FUNCTION_BLOCK PID_SAMPLE_COORDINATOR (* Experimental; offline checks only; native export/runtime pending *)
  (* Standard: 61499-2 *)
  (* Version 0.1, 2026-10-20, Guilherme *)
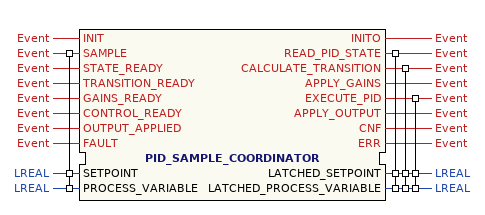
  EVENT_INPUT
    INIT;
    SAMPLE WITH SETPOINT, PROCESS_VARIABLE;
    STATE_READY;
    TRANSITION_READY;
    GAINS_READY;
    CONTROL_READY;
    OUTPUT_APPLIED;
    FAULT;
  END_EVENT
  EVENT_OUTPUT
    INITO;
    READ_PID_STATE WITH LATCHED_SETPOINT, LATCHED_PROCESS_VARIABLE;
    CALCULATE_TRANSITION WITH LATCHED_SETPOINT, LATCHED_PROCESS_VARIABLE;
    APPLY_GAINS;
    EXECUTE_PID WITH LATCHED_SETPOINT, LATCHED_PROCESS_VARIABLE;
    APPLY_OUTPUT;
    CNF;
    ERR;
  END_EVENT
  VAR_INPUT
    SETPOINT : LREAL;
    PROCESS_VARIABLE : LREAL;
  END_VAR
  VAR_OUTPUT
    LATCHED_SETPOINT : LREAL;
    LATCHED_PROCESS_VARIABLE : LREAL;
  END_VAR
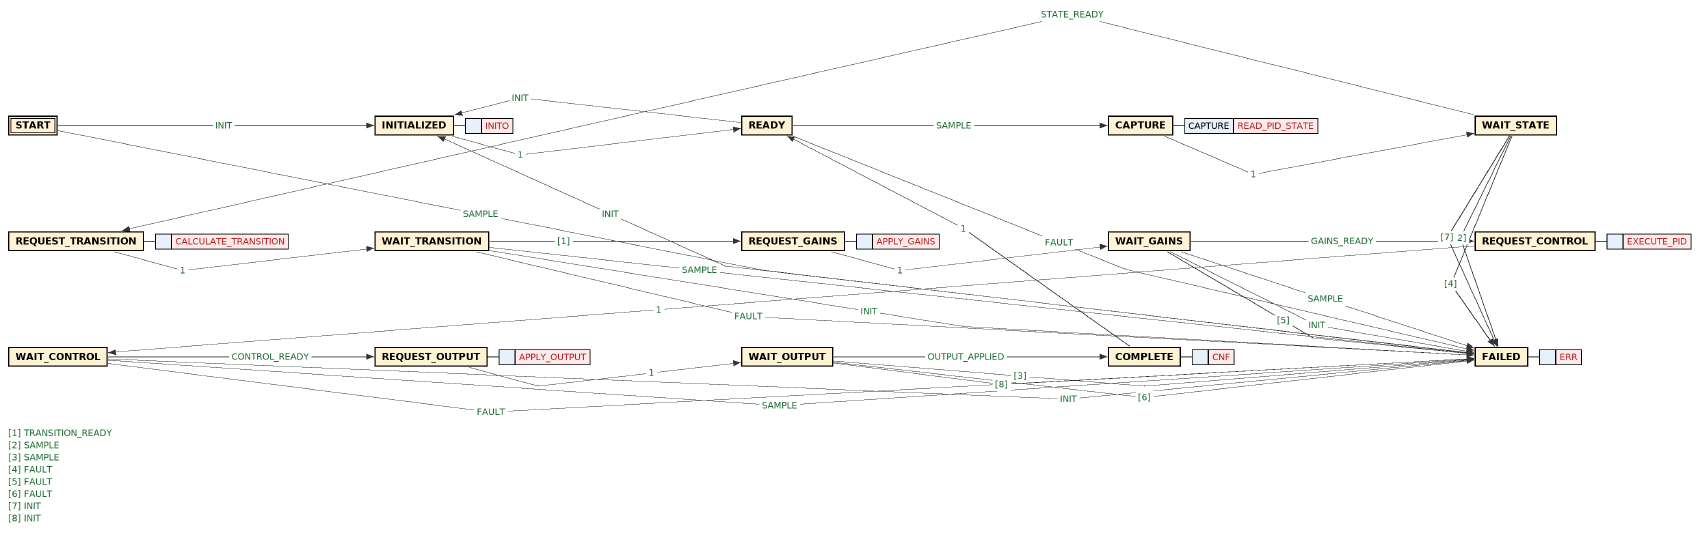
  EC_STATES
    START;
    INITIALIZED : -> INITO;
    READY;
    CAPTURE : CAPTURE -> READ_PID_STATE;
    WAIT_STATE;
    REQUEST_TRANSITION : -> CALCULATE_TRANSITION;
    WAIT_TRANSITION;
    REQUEST_GAINS : -> APPLY_GAINS;
    WAIT_GAINS;
    REQUEST_CONTROL : -> EXECUTE_PID;
    WAIT_CONTROL;
    REQUEST_OUTPUT : -> APPLY_OUTPUT;
    WAIT_OUTPUT;
    COMPLETE : -> CNF;
    FAILED : -> ERR;
  END_STATES
  EC_TRANSITIONS
    START TO INITIALIZED := INIT;
    INITIALIZED TO READY := 1;
    FAILED TO INITIALIZED := INIT;
    READY TO INITIALIZED := INIT;
    START TO FAILED := SAMPLE;
    READY TO CAPTURE := SAMPLE;
    CAPTURE TO WAIT_STATE := 1;
    WAIT_STATE TO REQUEST_TRANSITION := STATE_READY;
    REQUEST_TRANSITION TO WAIT_TRANSITION := 1;
    WAIT_STATE TO FAILED := SAMPLE;
    WAIT_STATE TO FAILED := INIT;
    WAIT_STATE TO FAILED := FAULT;
    WAIT_TRANSITION TO REQUEST_GAINS := TRANSITION_READY;
    REQUEST_GAINS TO WAIT_GAINS := 1;
    WAIT_TRANSITION TO FAILED := SAMPLE;
    WAIT_TRANSITION TO FAILED := INIT;
    WAIT_TRANSITION TO FAILED := FAULT;
    WAIT_GAINS TO REQUEST_CONTROL := GAINS_READY;
    REQUEST_CONTROL TO WAIT_CONTROL := 1;
    WAIT_GAINS TO FAILED := SAMPLE;
    WAIT_GAINS TO FAILED := INIT;
    WAIT_GAINS TO FAILED := FAULT;
    WAIT_CONTROL TO REQUEST_OUTPUT := CONTROL_READY;
    REQUEST_OUTPUT TO WAIT_OUTPUT := 1;
    WAIT_CONTROL TO FAILED := SAMPLE;
    WAIT_CONTROL TO FAILED := INIT;
    WAIT_CONTROL TO FAILED := FAULT;
    WAIT_OUTPUT TO COMPLETE := OUTPUT_APPLIED;
    COMPLETE TO READY := 1;
    WAIT_OUTPUT TO FAILED := SAMPLE;
    WAIT_OUTPUT TO FAILED := INIT;
    WAIT_OUTPUT TO FAILED := FAULT;
    READY TO FAILED := FAULT;
  END_TRANSITIONS
  ALGORITHM CAPTURE IN ST:
LATCHED_SETPOINT := SETPOINT;
LATCHED_PROCESS_VARIABLE := PROCESS_VARIABLE;
  END_ALGORITHM
END_FUNCTION_BLOCK
